FUNCTION_BLOCK Testing (* CAT Function Block Type *)
  (* Standard: 61499-2 *)
  (* Version 0.0, 11/20/2026, Schneider Electric, template *)
  PACKAGE Main;
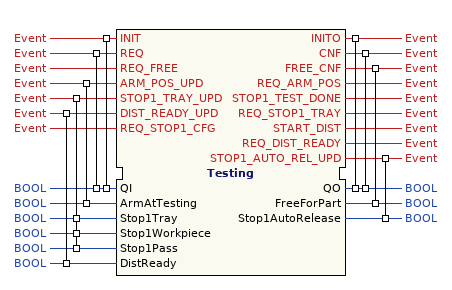
  EVENT_INPUT
    INIT WITH QI; (* Initialization Request *)
    REQ WITH QI; (* Normal Execution Request *)
    REQ_FREE; (* Request current downstream-free status *)
    ARM_POS_UPD WITH ArmAtTesting; (* Update Distribution swivel arm-at-Testing state *)
    STOP1_TRAY_UPD WITH Stop1Tray, Stop1Workpiece, Stop1Pass; (* Update Stop 1 tray and workpiece sensor states *)
    DIST_READY_UPD WITH DistReady; (* Update Distribution cycle ready state *)
    REQ_STOP1_CFG; (* Request current Stop 1 auto-release configuration from Conveyor on startup *)
  END_EVENT
  EVENT_OUTPUT
    INITO WITH QO; (* Initialization Confirm *)
    CNF WITH QO; (* Execution Confirmation *)
    FREE_CNF WITH FreeForPart; (* Downstream-free status changed *)
    REQ_ARM_POS; (* Request initial swivel arm position from Distribution on startup *)
    STOP1_TEST_DONE; (* Primary Station 1 Testing pass-complete notification to Conveyor Stop 1 *)
    REQ_STOP1_TRAY; (* Request initial Stop 1 tray/workpiece state from Conveyor *)
    START_DIST; (* Start Distribution AutoCycle programmatically *)
    REQ_DIST_READY; (* Request initial Distribution ready state *)
    STOP1_AUTO_REL_UPD WITH Stop1AutoRelease; (* Stop 1 auto-release enable update to Conveyor *)
  END_EVENT
  VAR_INPUT
    QI : BOOL; (* Input event qualifier *)
    ArmAtTesting : BOOL; (* TRUE when Distribution swivel arm is at Testing (3B2) *)
    Stop1Tray : BOOL; (* Tray present at Conveyor Stop 1 *)
    Stop1Workpiece : BOOL; (* Workpiece in Station 1 pocket at Stop 1 *)
    Stop1Pass : BOOL := FALSE; (* Stopper 1 pass-through or releasing state (TRUE=Down, FALSE=Up/Blocking) *)
    DistReady : BOOL := TRUE; (* TRUE when Distribution CycleSeq is Stopped or Completed (defaults TRUE standalone) *)
  END_VAR
  VAR_OUTPUT
    QO : BOOL; (* Output event qualifier *)
    FreeForPart : BOOL; (* TRUE when lift is lowered, ejector retracted, and no workpiece is present *)
    Stop1AutoRelease : BOOL; (* Effective Stop 1 auto-release enable (Auto S1 AND Auto-Rel) *)
  END_VAR
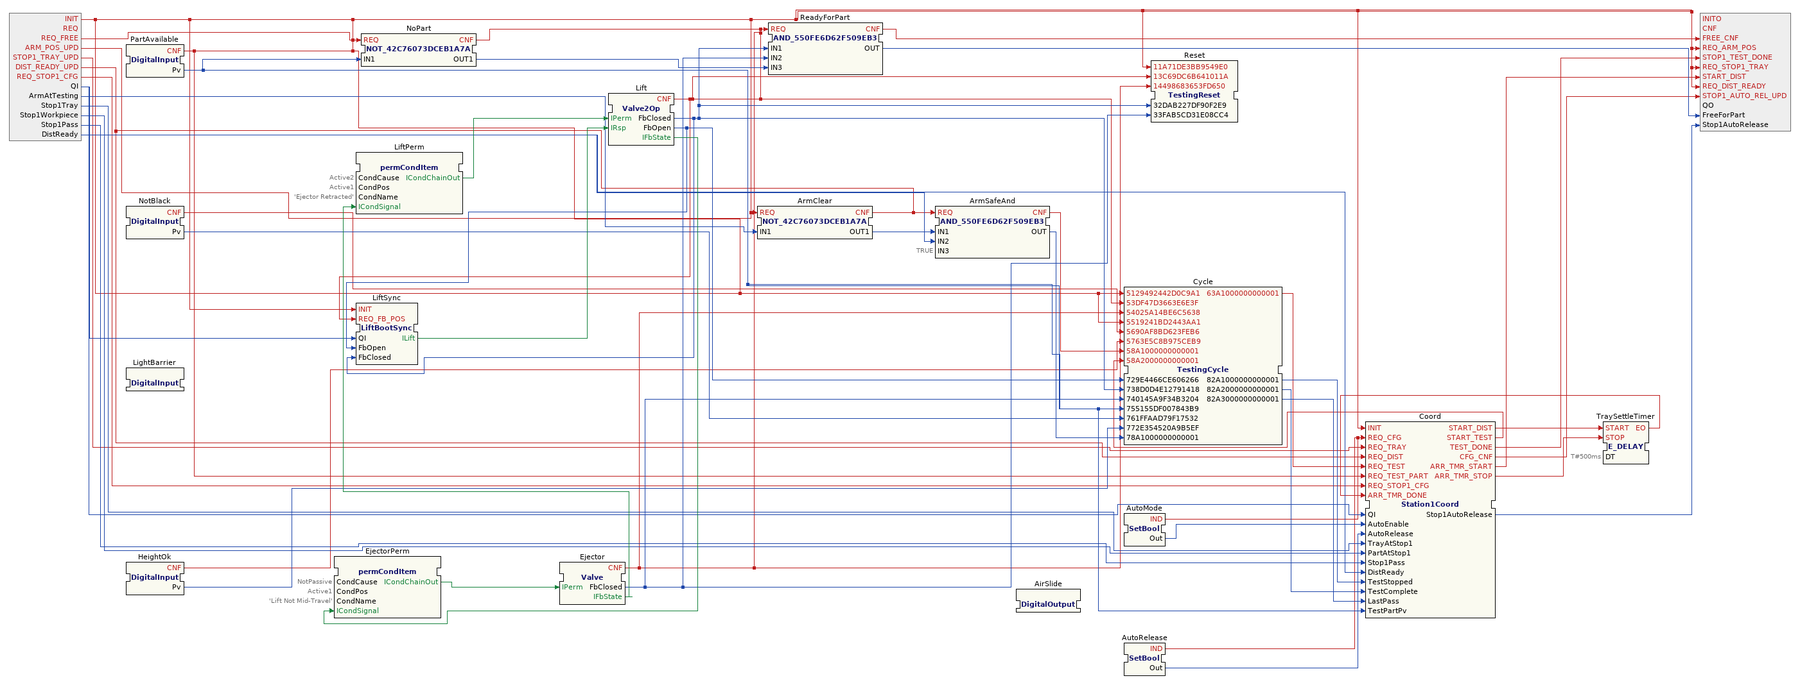
  FBS
    Lift : Valve2Op;
    Ejector : Valve;
    AirSlide : DigitalOutput;
    PartAvailable : DigitalInput;
    NotBlack : DigitalInput;
    LightBarrier : DigitalInput;
    HeightOk : DigitalInput;
    LiftPerm : permCondItem(CondCause := Active2, CondPos := Active1, CondName := 'Ejector Retracted');
    EjectorPerm : permCondItem(CondCause := NotPassive, CondPos := Active1, CondName := 'Lift Not Mid-Travel');
    Reset : TestingReset;
    Cycle : TestingCycle;
    NoPart : NOT_42C76073DCEB1A7A; {SET_ATTRIBUTE(Configuration.GenericFBType.InterfaceParams, Runtime.Standard#CNT:=1;OUT${CNT$}:BOOL)}
    ReadyForPart : AND_550FE6D62F509EB3; {SET_ATTRIBUTE(Configuration.GenericFBType.InterfaceParams, Runtime.Standard#CNT:=3;OUT:BOOL)}
    ArmClear : NOT_42C76073DCEB1A7A; {SET_ATTRIBUTE(Configuration.GenericFBType.InterfaceParams, Runtime.Standard#CNT:=1;OUT${CNT$}:BOOL)}
    AutoMode : SetBool;
    AutoRelease : SetBool;
    Coord : Station1Coord;
    TraySettleTimer : E_DELAY(DT := T#500ms);
    ArmSafeAnd : AND_550FE6D62F509EB3(IN3 := TRUE); {SET_ATTRIBUTE(Configuration.GenericFBType.InterfaceParams, Runtime.Standard#CNT:=3;OUT:BOOL)}
    LiftSync : LiftBootSync;
  END_FBS
  EVENT_CONNECTIONS
    INIT TO Reset.11A71DE3BB9549E0;
    INIT TO Cycle.5129492442D0C9A1;
    Lift.CNF TO Reset.13C69DC6B641011A;
    Ejector.CNF TO Reset.14498683653FD650;
    Lift.CNF TO Cycle.53DF47D3663E6E3F;
    Ejector.CNF TO Cycle.54025A14BE6C5638;
    PartAvailable.CNF TO Cycle.5519241BD2443AA1;
    NotBlack.CNF TO Cycle.5690AF8BD623FEB6;
    HeightOk.CNF TO Cycle.5763E5C8B975CEB9;
    INIT TO NoPart.REQ;
    REQ_FREE TO NoPart.REQ;
    PartAvailable.CNF TO NoPart.REQ;
    NoPart.CNF TO ReadyForPart.REQ;
    Lift.CNF TO ReadyForPart.REQ;
    Ejector.CNF TO ReadyForPart.REQ;
    ReadyForPart.CNF TO FREE_CNF;
    INIT TO ArmClear.REQ;
    INIT TO REQ_ARM_POS;
    ARM_POS_UPD TO ArmClear.REQ;
    ArmClear.CNF TO ArmSafeAnd.REQ;
    DIST_READY_UPD TO ArmSafeAnd.REQ;
    ArmSafeAnd.CNF TO Cycle.58A1000000000001;
    INIT TO LiftSync.INIT;
    Lift.CNF TO LiftSync.REQ_FB_POS;
    INIT TO Coord.INIT;
    INIT TO REQ_STOP1_TRAY;
    INIT TO REQ_DIST_READY;
    AutoMode.IND TO Coord.REQ_CFG;
    AutoRelease.IND TO Coord.REQ_CFG;
    STOP1_TRAY_UPD TO Coord.REQ_TRAY;
    DIST_READY_UPD TO Coord.REQ_DIST;
    Cycle.63A1000000000001 TO Coord.REQ_TEST;
    PartAvailable.CNF TO Coord.REQ_TEST_PART;
    REQ_STOP1_CFG TO Coord.REQ_STOP1_CFG;
    Coord.START_DIST TO START_DIST;
    Coord.START_TEST TO Cycle.58A2000000000001;
    Coord.TEST_DONE TO STOP1_TEST_DONE;
    Coord.CFG_CNF TO STOP1_AUTO_REL_UPD;
    Coord.ARR_TMR_START TO TraySettleTimer.START;
    Coord.ARR_TMR_STOP TO TraySettleTimer.STOP;
    TraySettleTimer.EO TO Coord.ARR_TMR_DONE;
  END_CONNECTIONS
  DATA_CONNECTIONS
    Lift.FbClosed TO Reset.32DAB227DF90F2E9;
    Ejector.FbClosed TO Reset.33FAB5CD31E08CC4;
    Lift.FbOpen TO Cycle.729E4466CE606266;
    Lift.FbClosed TO Cycle.738D0D4E12791418;
    Ejector.FbClosed TO Cycle.740145A9F34B3204;
    PartAvailable.Pv TO Cycle.755155DF007843B9;
    NotBlack.Pv TO Cycle.761FFAAD79F17532;
    HeightOk.Pv TO Cycle.772E354520A9B5EF;
    PartAvailable.Pv TO NoPart.IN1;
    Lift.FbClosed TO ReadyForPart.IN1;
    Ejector.FbClosed TO ReadyForPart.IN2;
    NoPart.OUT1 TO ReadyForPart.IN3;
    ReadyForPart.OUT TO FreeForPart;
    ArmAtTesting TO ArmClear.IN1;
    ArmClear.OUT1 TO ArmSafeAnd.IN1;
    DistReady TO ArmSafeAnd.IN2;
    ArmSafeAnd.OUT TO Cycle.78A1000000000001;
    QI TO LiftSync.QI;
    Lift.FbOpen TO LiftSync.FbOpen;
    Lift.FbClosed TO LiftSync.FbClosed;
    QI TO Coord.QI;
    AutoMode.Out TO Coord.AutoEnable;
    AutoRelease.Out TO Coord.AutoRelease;
    Stop1Tray TO Coord.TrayAtStop1;
    Stop1Workpiece TO Coord.PartAtStop1;
    Stop1Pass TO Coord.Stop1Pass;
    DistReady TO Coord.DistReady;
    Cycle.82A1000000000001 TO Coord.TestStopped;
    Cycle.82A2000000000001 TO Coord.TestComplete;
    Cycle.82A3000000000001 TO Coord.LastPass;
    PartAvailable.Pv TO Coord.TestPartPv;
    Coord.Stop1AutoRelease TO Stop1AutoRelease;
  END_CONNECTIONS
  ADAPTER_CONNECTIONS
    Ejector.IFbState TO LiftPerm.ICondSignal;
    LiftPerm.ICondChainOut TO Lift.IPerm;
    Lift.IFbState TO EjectorPerm.ICondSignal;
    EjectorPerm.ICondChainOut TO Ejector.IPerm;
    LiftSync.ILift TO Lift.IRsp;
  END_CONNECTIONS
END_FUNCTION_BLOCK
